{attribute 'qualified_only'}
{attribute 'strict'}
{attribute 'to_string'}
TYPE E_Dint :
(
	eOptionA := 0,
	eOptionB,
	eOptionC
) DINT;
END_TYPE

(* stored: Version 1.1.0.1, ProductVersion 3.1.4026.19
   DUT E_Dint: Id {77a05564-7940-46a5-9f6f-1110d53014ec} *)
